// TIA Portal V19 export
DATA_BLOCK "TIMER_DB_3"   // DB17
// stored: InstanceOfName TIMER, InstanceOfType FB
"TIMER"
   // VAR_INPUT
   //    START_TIMER : Bool;
   //    HR_SET : Int;
   //    MIN_SET : Int;
   //    SEC_SET : Int;
   //    RESET_TIMER : Bool;
   // END_VAR
   // VAR_OUTPUT
   //    SEC : Int;
   //    MIN : Int;
   //    HR : Int;
   //    TIMER_DONE { ExternalAccessible := 'False'; ExternalVisible := 'False'; ExternalWritable := 'False'} : Bool;
   // END_VAR
   // VAR
   //    P_TRIG1 : Bool;
   //    P_TRIG2 : Bool;
   //    P_TRIG3 : Bool;
   // END_VAR
BEGIN
END_DATA_BLOCK
